Fanuc KAREL source: kt00551.KL

-- PROVISIONAL review KL for V770-1; original PC SHA256 4a041cfdb72b1b117e8f084b83babfb86bc3c2d5533c5ab62d4ee6347325de46
-- Incomplete behavior may be omitted. Consult companion uncertainty JSON. Do not deploy.
PROGRAM KT00551
%NOLOCKGROUP
-- UNRESOLVED_DECL P1 type=000199
-- UNRESOLVED_DECL P2 type=000199
-- UNRESOLVED_DECL OUT type=000106
BEGIN
  -- UNRESOLVED_PC offsets 5-44; opcodes 49,7E,49,7E,60,7E,4A
  -- UNRESOLVED_PC offsets 49-53; opcodes 7F
END KT00551
